(* IEC 61131-3 sources: trust-platform/crates/trust-runtime/tests/fixtures/control_pid/src, 10 files *)

(* ---- advanced_control_tests.st ---- *)
USING Control;

TEST_PROGRAM control_smith_predictor_models_delay_and_anchors_prediction_to_measurement
VAR
    Predictor : SmithPredictorFOPDT;
    Parameters : SmithPredictorParameters;
    State : SmithPredictorInitialState;
    Input : SmithPredictorInput;
    Output : SmithPredictorOutput;
    Accepted : BOOL;
END_VAR
Parameters.ProcessGain := LREAL#2.0;
Parameters.TimeConstant := LREAL#1.0;
Parameters.DeadTime := LREAL#1.0;
Parameters.OperatingOutput := LREAL#10.0;
Parameters.MaximumCorrection := LREAL#0.5;
Accepted := Predictor.Configure(Parameters := Parameters);
ASSERT_TRUE(Accepted);
State.ModelOutput := LREAL#10.0;
State.ProcessValue := LREAL#10.0;
Predictor.Initialize(State := State);
Input.ManipulatedValue := LREAL#1.0;
Input.ProcessValue := LREAL#10.0;
Input.CycleTime := LREAL#0.5;
Input.Enabled := TRUE;
Output := Predictor.Update(Input := Input);
ASSERT_TRUE(Output.Active);
ASSERT_TRUE(Output.HistoryComplete);
ASSERT_NEAR(EXPECTED := LREAL#10.8, ACTUAL := Output.DelayFreeModel, DELTA := LREAL#1.0e-12);
ASSERT_NEAR(EXPECTED := LREAL#10.0, ACTUAL := Output.DelayedModel, DELTA := LREAL#1.0e-12);
ASSERT_NEAR(EXPECTED := LREAL#10.8, ACTUAL := Output.PredictedProcessValue, DELTA := LREAL#1.0e-12);

Input.ProcessValue := LREAL#12.0;
Output := Predictor.Update(Input := Input);
ASSERT_NEAR(EXPECTED := LREAL#0.5, ACTUAL := Output.Correction, DELTA := LREAL#1.0e-12);
ASSERT_NEAR(EXPECTED := LREAL#11.78, ACTUAL := Output.PredictedProcessValue, DELTA := LREAL#1.0e-12);

Input.Enabled := FALSE;
Input.ProcessValue := LREAL#9.25;
Output := Predictor.Update(Input := Input);
ASSERT_FALSE(Output.Active);
ASSERT_NEAR(EXPECTED := LREAL#9.25, ACTUAL := Output.PredictedProcessValue, DELTA := LREAL#1.0e-12);

Parameters.TimeConstant := LREAL#0.0;
Accepted := Predictor.Configure(Parameters := Parameters);
ASSERT_FALSE(Accepted);
END_TEST_PROGRAM

TEST_PROGRAM control_pid_form_conversion_is_explicit_reversible_and_fail_closed
VAR
    Input : PIDFormParameters;
    Result : PIDFormConversionResult;
    Parallel : PIDFormParameters;
END_VAR

Input.Form := PIDParameterForm#Ideal;
Input.Proportional := LREAL#2.0;
Input.Integral := LREAL#10.0;
Input.Derivative := LREAL#0.5;
Result := ConvertPIDForm(Input := Input, Target := PIDParameterForm#Parallel);
ASSERT_TRUE(Result.Status = PIDFormConversionStatus#Valid);
ASSERT_NEAR(EXPECTED := LREAL#2.0, ACTUAL := Result.Parameters.Proportional, DELTA := LREAL#1.0e-12);
ASSERT_NEAR(EXPECTED := LREAL#0.2, ACTUAL := Result.Parameters.Integral, DELTA := LREAL#1.0e-12);
ASSERT_NEAR(EXPECTED := LREAL#1.0, ACTUAL := Result.Parameters.Derivative, DELTA := LREAL#1.0e-12);

Input.Form := PIDParameterForm#Series;
Result := ConvertPIDForm(Input := Input, Target := PIDParameterForm#Parallel);
ASSERT_TRUE(Result.Status = PIDFormConversionStatus#Valid);
ASSERT_NEAR(EXPECTED := LREAL#2.1, ACTUAL := Result.Parameters.Proportional, DELTA := LREAL#1.0e-12);
ASSERT_NEAR(EXPECTED := LREAL#0.2, ACTUAL := Result.Parameters.Integral, DELTA := LREAL#1.0e-12);
ASSERT_NEAR(EXPECTED := LREAL#1.0, ACTUAL := Result.Parameters.Derivative, DELTA := LREAL#1.0e-12);
Parallel := Result.Parameters;
Result := ConvertPIDForm(Input := Parallel, Target := PIDParameterForm#Series);
ASSERT_TRUE(Result.Status = PIDFormConversionStatus#Valid);
ASSERT_NEAR(EXPECTED := LREAL#2.0, ACTUAL := Result.Parameters.Proportional, DELTA := LREAL#1.0e-12);
ASSERT_NEAR(EXPECTED := LREAL#10.0, ACTUAL := Result.Parameters.Integral, DELTA := LREAL#1.0e-12);
ASSERT_NEAR(EXPECTED := LREAL#0.5, ACTUAL := Result.Parameters.Derivative, DELTA := LREAL#1.0e-12);

Parallel.Form := PIDParameterForm#Parallel;
Parallel.Proportional := LREAL#-2.0;
Parallel.Integral := LREAL#-0.2;
Parallel.Derivative := LREAL#-1.0;
Result := ConvertPIDForm(Input := Parallel, Target := PIDParameterForm#Ideal);
ASSERT_TRUE(Result.Status = PIDFormConversionStatus#Valid);
ASSERT_NEAR(EXPECTED := LREAL#-2.0, ACTUAL := Result.Parameters.Proportional, DELTA := LREAL#1.0e-12);
ASSERT_NEAR(EXPECTED := LREAL#10.0, ACTUAL := Result.Parameters.Integral, DELTA := LREAL#1.0e-12);
ASSERT_NEAR(EXPECTED := LREAL#0.5, ACTUAL := Result.Parameters.Derivative, DELTA := LREAL#1.0e-12);

Result := ConvertPIDForm(Input := Parallel, Target := PIDParameterForm#Parallel);
ASSERT_TRUE(Result.Status = PIDFormConversionStatus#Valid);
ASSERT_NEAR(EXPECTED := Parallel.Proportional, ACTUAL := Result.Parameters.Proportional, DELTA := LREAL#1.0e-12);

Input.Form := PIDParameterForm#Ideal;
Input.Proportional := LREAL#2.0;
Input.Integral := LREAL#0.0;
Input.Derivative := LREAL#0.5;
Result := ConvertPIDForm(Input := Input, Target := PIDParameterForm#Parallel);
ASSERT_TRUE(Result.Status = PIDFormConversionStatus#InvalidDomain);

Parallel.Form := PIDParameterForm#Parallel;
Parallel.Proportional := LREAL#1.0;
Parallel.Integral := LREAL#1.0;
Parallel.Derivative := LREAL#1.0;
Result := ConvertPIDForm(Input := Parallel, Target := PIDParameterForm#Series);
ASSERT_TRUE(Result.Status = PIDFormConversionStatus#NonRepresentable);
END_TEST_PROGRAM

TEST_PROGRAM control_smith_predictor_initialization_sets_the_correction_from_the_measurement
VAR
    Predictor : SmithPredictorFOPDT;
    State : SmithPredictorInitialState;
    Input : SmithPredictorInput;
    Output : SmithPredictorOutput;
END_VAR
(* Spec 37 §2.3: Initialize sets the initial correction from ProcessValue - ModelOutput. Before
   configuration no model interval runs, so the update reports that correction while it returns
   the measurement. *)
State.ModelOutput := LREAL#10.0;
State.ProcessValue := LREAL#12.0;
Predictor.Initialize(State := State);
Input.ProcessValue := LREAL#12.0;
Input.CycleTime := LREAL#0.5;
Input.Enabled := TRUE;
Output := Predictor.Update(Input := Input);
ASSERT_FALSE(Output.Active);
ASSERT_NEAR(EXPECTED := LREAL#12.0, ACTUAL := Output.PredictedProcessValue, DELTA := LREAL#1.0e-12);
ASSERT_NEAR(EXPECTED := LREAL#2.0, ACTUAL := Output.Correction, DELTA := LREAL#1.0e-12);
END_TEST_PROGRAM

TEST_PROGRAM control_smith_predictor_zero_delay_reduces_to_measurement
VAR
    Predictor : SmithPredictorFOPDT;
    Parameters : SmithPredictorParameters;
    State : SmithPredictorInitialState;
    Input : SmithPredictorInput;
    Output : SmithPredictorOutput;
END_VAR
Parameters.ProcessGain := LREAL#1.0;
Parameters.TimeConstant := LREAL#2.0;
Parameters.DeadTime := LREAL#0.0;
ASSERT_TRUE(Predictor.Configure(Parameters := Parameters));
Predictor.Initialize(State := State);
Input.ManipulatedValue := LREAL#4.0;
Input.ProcessValue := LREAL#7.25;
Input.CycleTime := LREAL#0.1;
Input.Enabled := TRUE;
Output := Predictor.Update(Input := Input);
ASSERT_NEAR(EXPECTED := LREAL#7.25, ACTUAL := Output.PredictedProcessValue, DELTA := LREAL#1.0e-12);
END_TEST_PROGRAM

TEST_PROGRAM control_pid_gain_scheduler_interpolates_tuning_and_preserves_common_policy
VAR
    Scheduler : PIDGainScheduler;
    Parameters : PIDGainScheduleParameters;
    Output : PIDGainScheduleOutput;
    Accepted : BOOL;
END_VAR
Parameters.PointCount := DINT#3;
Parameters.Points[0].OperatingPoint := LREAL#0.0;
Parameters.Points[0].Tuning.ProportionalGain := LREAL#1.0;
Parameters.Points[0].Tuning.IntegralGain := LREAL#0.1;
Parameters.Points[0].Tuning.DerivativeGain := LREAL#0.2;
Parameters.Points[0].Tuning.ProportionalSetpointWeight := LREAL#0.3;
Parameters.Points[0].Tuning.DerivativeSetpointWeight := LREAL#0.4;
Parameters.Points[0].Tuning.TrackingTime := LREAL#1.0;
Parameters.Points[1].OperatingPoint := LREAL#10.0;
Parameters.Points[1].Tuning.ProportionalGain := LREAL#2.0;
Parameters.Points[1].Tuning.IntegralGain := LREAL#0.2;
Parameters.Points[1].Tuning.DerivativeGain := LREAL#0.4;
Parameters.Points[1].Tuning.ProportionalSetpointWeight := LREAL#0.5;
Parameters.Points[1].Tuning.DerivativeSetpointWeight := LREAL#0.6;
Parameters.Points[1].Tuning.TrackingTime := LREAL#2.0;
Parameters.Points[2].OperatingPoint := LREAL#20.0;
Parameters.Points[2].Tuning.ProportionalGain := LREAL#4.0;
Parameters.Points[2].Tuning.IntegralGain := LREAL#0.4;
Parameters.Points[2].Tuning.DerivativeGain := LREAL#0.8;
Parameters.Points[2].Tuning.ProportionalSetpointWeight := LREAL#0.7;
Parameters.Points[2].Tuning.DerivativeSetpointWeight := LREAL#0.8;
Parameters.Points[2].Tuning.TrackingTime := LREAL#4.0;
Parameters.CommonParameters.Bias := LREAL#12.0;
Parameters.CommonParameters.OutputMinimum := LREAL#0.0;
Parameters.CommonParameters.OutputMaximum := LREAL#100.0;
Parameters.CommonParameters.RateMinimum := LREAL#-5.0;
Parameters.CommonParameters.RateMaximum := LREAL#7.0;
Parameters.CommonParameters.AntiWindup := PIDAntiWindup#Combined;
Accepted := Scheduler.Configure(Parameters := Parameters);
ASSERT_TRUE(Accepted);
Scheduler.Initialize(OperatingPoint := LREAL#5.0);
Output := Scheduler.Update(OperatingPoint := LREAL#5.0, CycleTime := LREAL#0.1);
ASSERT_TRUE(Output.Valid);
ASSERT_FALSE(Output.Clamped);
ASSERT_TRUE(Output.LowerIndex = DINT#0);
ASSERT_TRUE(Output.UpperIndex = DINT#1);
ASSERT_NEAR(EXPECTED := LREAL#0.5, ACTUAL := Output.Fraction, DELTA := LREAL#1.0e-12);
ASSERT_NEAR(EXPECTED := LREAL#1.5, ACTUAL := Output.Parameters.ProportionalGain, DELTA := LREAL#1.0e-12);
ASSERT_NEAR(EXPECTED := LREAL#0.15, ACTUAL := Output.Parameters.IntegralGain, DELTA := LREAL#1.0e-12);
ASSERT_NEAR(EXPECTED := LREAL#0.3, ACTUAL := Output.Parameters.DerivativeGain, DELTA := LREAL#1.0e-12);
ASSERT_NEAR(EXPECTED := LREAL#0.4, ACTUAL := Output.Parameters.ProportionalSetpointWeight, DELTA := LREAL#1.0e-12);
ASSERT_NEAR(EXPECTED := LREAL#0.5, ACTUAL := Output.Parameters.DerivativeSetpointWeight, DELTA := LREAL#1.0e-12);
ASSERT_NEAR(EXPECTED := LREAL#1.5, ACTUAL := Output.Parameters.TrackingTime, DELTA := LREAL#1.0e-12);
ASSERT_NEAR(EXPECTED := LREAL#12.0, ACTUAL := Output.Parameters.Bias, DELTA := LREAL#1.0e-12);
ASSERT_NEAR(EXPECTED := LREAL#100.0, ACTUAL := Output.Parameters.OutputMaximum, DELTA := LREAL#1.0e-12);
ASSERT_TRUE(Output.Parameters.AntiWindup = PIDAntiWindup#Combined);

Output := Scheduler.Update(OperatingPoint := LREAL#-5.0, CycleTime := LREAL#0.1);
ASSERT_TRUE(Output.Clamped);
ASSERT_NEAR(EXPECTED := LREAL#1.0, ACTUAL := Output.Parameters.ProportionalGain, DELTA := LREAL#1.0e-12);

Parameters.Points[1].OperatingPoint := LREAL#0.0;
Accepted := Scheduler.Configure(Parameters := Parameters);
ASSERT_FALSE(Accepted);
Output := Scheduler.Update(OperatingPoint := LREAL#15.0, CycleTime := LREAL#0.1);
ASSERT_NEAR(EXPECTED := LREAL#3.0, ACTUAL := Output.Parameters.ProportionalGain, DELTA := LREAL#1.0e-12);
END_TEST_PROGRAM

TEST_PROGRAM control_pid_gain_scheduler_filters_the_operating_point
VAR
    Scheduler : PIDGainScheduler;
    Parameters : PIDGainScheduleParameters;
    Output : PIDGainScheduleOutput;
END_VAR
Parameters.PointCount := DINT#2;
Parameters.Points[0].OperatingPoint := LREAL#0.0;
Parameters.Points[0].Tuning.ProportionalGain := LREAL#1.0;
Parameters.Points[0].Tuning.TrackingTime := LREAL#1.0;
Parameters.Points[1].OperatingPoint := LREAL#10.0;
Parameters.Points[1].Tuning.ProportionalGain := LREAL#3.0;
Parameters.Points[1].Tuning.TrackingTime := LREAL#1.0;
Parameters.CommonParameters.OutputMinimum := LREAL#-100.0;
Parameters.CommonParameters.OutputMaximum := LREAL#100.0;
Parameters.CommonParameters.RateMinimum := LREAL#-100.0;
Parameters.CommonParameters.RateMaximum := LREAL#100.0;
Parameters.FilterTimeConstant := LREAL#1.0;
ASSERT_TRUE(Scheduler.Configure(Parameters := Parameters));
Scheduler.Initialize(OperatingPoint := LREAL#0.0);
Output := Scheduler.Update(OperatingPoint := LREAL#10.0, CycleTime := LREAL#1.0);
ASSERT_NEAR(EXPECTED := LREAL#5.0, ACTUAL := Output.FilteredOperatingPoint, DELTA := LREAL#1.0e-12);
ASSERT_NEAR(EXPECTED := LREAL#2.0, ACTUAL := Output.Parameters.ProportionalGain, DELTA := LREAL#1.0e-12);
END_TEST_PROGRAM

TEST_PROGRAM control_static_decoupler_maps_and_recovers_two_channel_commands
VAR
    Decoupler : StaticDecoupler2x2;
    Parameters : StaticDecoupler2x2Parameters;
    VirtualCommand : ControlVector2;
    ActuatorCommand : ControlVector2;
    Recovered : ControlVector2;
    Status : StaticDecoupler2x2Status;
    Accepted : BOOL;
END_VAR
VirtualCommand.First := LREAL#3.0;
ActuatorCommand := Decoupler.ToActuators(VirtualCommand := VirtualCommand);
ASSERT_NEAR(EXPECTED := LREAL#0.0, ACTUAL := ActuatorCommand.First, DELTA := LREAL#1.0e-12);
ASSERT_NEAR(EXPECTED := LREAL#0.0, ACTUAL := ActuatorCommand.Second, DELTA := LREAL#1.0e-12);

Parameters.GainMatrix.G11 := LREAL#2.0;
Parameters.GainMatrix.G12 := LREAL#1.0;
Parameters.GainMatrix.G21 := LREAL#1.0;
Parameters.GainMatrix.G22 := LREAL#2.0;
Parameters.ActuatorBias.First := LREAL#10.0;
Parameters.ActuatorBias.Second := LREAL#20.0;
Parameters.SingularityTolerance := LREAL#1.0e-9;
Accepted := Decoupler.Configure(Parameters := Parameters);
ASSERT_TRUE(Accepted);
Status := Decoupler.Snapshot();
ASSERT_TRUE(Status.Configured);
ASSERT_NEAR(EXPECTED := LREAL#3.0, ACTUAL := Status.Determinant, DELTA := LREAL#1.0e-12);
ActuatorCommand := Decoupler.ToActuators(VirtualCommand := VirtualCommand);
ASSERT_NEAR(EXPECTED := LREAL#12.0, ACTUAL := ActuatorCommand.First, DELTA := LREAL#1.0e-12);
ASSERT_NEAR(EXPECTED := LREAL#19.0, ACTUAL := ActuatorCommand.Second, DELTA := LREAL#1.0e-12);
Recovered := Decoupler.ToVirtual(ActuatorCommand := ActuatorCommand);
ASSERT_NEAR(EXPECTED := LREAL#3.0, ACTUAL := Recovered.First, DELTA := LREAL#1.0e-12);
ASSERT_NEAR(EXPECTED := LREAL#0.0, ACTUAL := Recovered.Second, DELTA := LREAL#1.0e-12);

Parameters.GainMatrix.G11 := LREAL#1000000.0;
Parameters.GainMatrix.G12 := LREAL#1000000.0;
Parameters.GainMatrix.G21 := LREAL#1000000.0;
Parameters.GainMatrix.G22 := LREAL#1000000.01;
Parameters.SingularityTolerance := LREAL#1.0e-6;
Accepted := Decoupler.Configure(Parameters := Parameters);
ASSERT_FALSE(Accepted);
ActuatorCommand := Decoupler.ToActuators(VirtualCommand := VirtualCommand);
ASSERT_NEAR(EXPECTED := LREAL#12.0, ACTUAL := ActuatorCommand.First, DELTA := LREAL#1.0e-12);
ASSERT_NEAR(EXPECTED := LREAL#19.0, ACTUAL := ActuatorCommand.Second, DELTA := LREAL#1.0e-12);

Parameters.GainMatrix.G11 := LREAL#1.0;
Parameters.GainMatrix.G12 := LREAL#2.0;
Parameters.GainMatrix.G21 := LREAL#2.0;
Parameters.GainMatrix.G22 := LREAL#4.0;
Accepted := Decoupler.Configure(Parameters := Parameters);
ASSERT_FALSE(Accepted);
ActuatorCommand := Decoupler.ToActuators(VirtualCommand := VirtualCommand);
ASSERT_NEAR(EXPECTED := LREAL#12.0, ACTUAL := ActuatorCommand.First, DELTA := LREAL#1.0e-12);
ASSERT_NEAR(EXPECTED := LREAL#19.0, ACTUAL := ActuatorCommand.Second, DELTA := LREAL#1.0e-12);
END_TEST_PROGRAM

(* ---- antiwindup_tests.st ---- *)
USING Control;

TEST_PROGRAM control_pid_back_calculation_and_clamping_retain_distinct_nominal_states
VAR
    BackCalculationController : PID;
    ClampingController : PID;
    Parameters : PIDParameters;
    InitialState : PIDInitialState;
    Input : PIDInput;
    Output : LREAL;
END_VAR

Parameters.IntegralGain := LREAL#4.0;
Parameters.OutputMinimum := LREAL#0.0;
Parameters.OutputMaximum := LREAL#3.0;
Parameters.RateMinimum := LREAL#-1000.0;
Parameters.RateMaximum := LREAL#1000.0;
Parameters.TrackingTime := LREAL#2.0;
BackCalculationController.Configure(Parameters := Parameters);
BackCalculationController.Initialize(State := InitialState);

Input.Setpoint := LREAL#1.0;
Input.CycleTime := LREAL#1.0;
Output := BackCalculationController.Update(Input := Input);
ASSERT_NEAR(EXPECTED := LREAL#3.0, ACTUAL := Output, DELTA := LREAL#3.0e-12);
Input.Setpoint := LREAL#-0.125;
Output := BackCalculationController.Update(Input := Input);
ASSERT_NEAR(EXPECTED := LREAL#3.0, ACTUAL := Output, DELTA := LREAL#3.0e-12);

Parameters.TrackingTime := LREAL#1.0;
ClampingController.Configure(Parameters := Parameters);
ClampingController.Initialize(State := InitialState);
Input.Setpoint := LREAL#1.0;
Output := ClampingController.Update(Input := Input);
ASSERT_NEAR(EXPECTED := LREAL#3.0, ACTUAL := Output, DELTA := LREAL#3.0e-12);
Input.Setpoint := LREAL#-0.125;
Output := ClampingController.Update(Input := Input);
ASSERT_NEAR(EXPECTED := LREAL#2.5, ACTUAL := Output, DELTA := LREAL#2.5e-12);
END_TEST_PROGRAM

TEST_PROGRAM control_pid_combined_anti_windup_allows_integration_away_from_saturation
VAR
    Controller : PID;
    Parameters : PIDParameters;
    InitialState : PIDInitialState;
    Input : PIDInput;
    Output : LREAL;
END_VAR

Parameters.IntegralGain := LREAL#1.0;
Parameters.OutputMinimum := LREAL#0.0;
Parameters.OutputMaximum := LREAL#3.0;
Parameters.RateMinimum := LREAL#-1000.0;
Parameters.RateMaximum := LREAL#1000.0;
Parameters.TrackingTime := LREAL#2.0;
Parameters.AntiWindup := PIDAntiWindup#Combined;
InitialState.NominalOutput := LREAL#4.0;
InitialState.SaturatedOutput := LREAL#3.0;
Controller.Configure(Parameters := Parameters);
Controller.Initialize(State := InitialState);

Input.Setpoint := LREAL#1.0;
Input.CycleTime := LREAL#1.0;
Output := Controller.Update(Input := Input);
ASSERT_NEAR(EXPECTED := LREAL#3.0, ACTUAL := Output, DELTA := LREAL#3.0e-12);

Input.Setpoint := LREAL#-0.75;
Output := Controller.Update(Input := Input);
ASSERT_NEAR(EXPECTED := LREAL#2.75, ACTUAL := Output, DELTA := LREAL#2.75e-12);
END_TEST_PROGRAM

(* ---- configuration_tests.st ---- *)
(* Specification 45 sections 2.4/2.5 and 3.2/3.3: complete value-copy configuration,
   retained histories, and initialization without an update. *)
USING Control;

TEST_PROGRAM control_pid_configuration_copies_parameters_and_preserves_every_history
VAR
    Controller : PID;
    Parameters : PIDParameters;
    AcceptedParameters : PIDParameters;
    InitialState : PIDInitialState;
    ZeroState : PIDInitialState;
    Observed : PIDInitialState;
    Input : PIDInput;
    Output : LREAL;
END_VAR

InitialState.Setpoint := LREAL#10.0;
InitialState.SetpointRate := LREAL#2.0;
InitialState.ProcessValue := LREAL#8.0;
InitialState.ProcessValueRate := LREAL#-1.0;
InitialState.FeedForward := LREAL#3.0;
InitialState.NominalOutput := LREAL#20.0;
InitialState.SaturatedOutput := LREAL#19.0;
Parameters.OutputMinimum := LREAL#-100.0;
Parameters.OutputMaximum := LREAL#100.0;
Parameters.RateMinimum := LREAL#-1000.0;
Parameters.RateMaximum := LREAL#1000.0;
Parameters.TrackingTime := LREAL#1.0;
Controller.Configure(Parameters := Parameters);
Controller.Initialize(State := InitialState);
Observed := Controller.GetState();
ASSERT_NEAR(EXPECTED := LREAL#10.0, ACTUAL := Observed.Setpoint, DELTA := LREAL#1.0e-12);
ASSERT_NEAR(EXPECTED := LREAL#2.0, ACTUAL := Observed.SetpointRate, DELTA := LREAL#1.0e-12);
ASSERT_NEAR(EXPECTED := LREAL#8.0, ACTUAL := Observed.ProcessValue, DELTA := LREAL#1.0e-12);
ASSERT_NEAR(EXPECTED := LREAL#-1.0, ACTUAL := Observed.ProcessValueRate, DELTA := LREAL#1.0e-12);
ASSERT_NEAR(EXPECTED := LREAL#3.0, ACTUAL := Observed.FeedForward, DELTA := LREAL#1.0e-12);
ASSERT_NEAR(EXPECTED := LREAL#20.0, ACTUAL := Observed.NominalOutput, DELTA := LREAL#1.0e-12);
ASSERT_NEAR(EXPECTED := LREAL#19.0, ACTUAL := Observed.SaturatedOutput, DELTA := LREAL#1.0e-12);

Parameters.ProportionalGain := LREAL#2.0;
Parameters.IntegralGain := LREAL#0.5;
Parameters.DerivativeGain := LREAL#0.25;
Parameters.ProportionalSetpointWeight := LREAL#0.4;
Parameters.DerivativeSetpointWeight := LREAL#0.3;
Parameters.Bias := LREAL#7.0;
Parameters.OutputMinimum := LREAL#-30.0;
Parameters.OutputMaximum := LREAL#40.0;
Parameters.RateMinimum := LREAL#-4.0;
Parameters.RateMaximum := LREAL#6.0;
Parameters.TrackingTime := LREAL#2.0;
Parameters.AntiWindup := PIDAntiWindup#Combined;
Controller.Configure(Parameters := Parameters);
Observed := Controller.GetState();
ASSERT_NEAR(EXPECTED := LREAL#10.0, ACTUAL := Observed.Setpoint, DELTA := LREAL#1.0e-12);
ASSERT_NEAR(EXPECTED := LREAL#2.0, ACTUAL := Observed.SetpointRate, DELTA := LREAL#1.0e-12);
ASSERT_NEAR(EXPECTED := LREAL#8.0, ACTUAL := Observed.ProcessValue, DELTA := LREAL#1.0e-12);
ASSERT_NEAR(EXPECTED := LREAL#-1.0, ACTUAL := Observed.ProcessValueRate, DELTA := LREAL#1.0e-12);
ASSERT_NEAR(EXPECTED := LREAL#3.0, ACTUAL := Observed.FeedForward, DELTA := LREAL#1.0e-12);
ASSERT_NEAR(EXPECTED := LREAL#20.0, ACTUAL := Observed.NominalOutput, DELTA := LREAL#1.0e-12);
ASSERT_NEAR(EXPECTED := LREAL#19.0, ACTUAL := Observed.SaturatedOutput, DELTA := LREAL#1.0e-12);

(* Mutating the caller's record after Configure cannot alter the accepted copy. *)
AcceptedParameters := Parameters;
Parameters.ProportionalGain := LREAL#100.0;
Parameters.IntegralGain := LREAL#0.0;
Parameters.DerivativeGain := LREAL#0.0;
Parameters.ProportionalSetpointWeight := LREAL#1.0;
Parameters.DerivativeSetpointWeight := LREAL#1.0;
Parameters.Bias := LREAL#-10.0;
Parameters.OutputMinimum := LREAL#-100.0;
Parameters.OutputMaximum := LREAL#100.0;
Parameters.RateMinimum := LREAL#-1000.0;
Parameters.RateMaximum := LREAL#1000.0;
Parameters.TrackingTime := LREAL#10.0;
Parameters.AntiWindup := PIDAntiWindup#BackCalculation;

Input.Setpoint := LREAL#12.0;
Input.ProcessValue := LREAL#9.0;
Input.FeedForward := LREAL#5.0;
Input.CycleTime := LREAL#0.5;
Output := Controller.Update(Input := Input);
(* 20 - 0.4 + 0.75 - 0.6 + 2 = 21.75; rate interval is [17,22]. *)
ASSERT_NEAR(EXPECTED := LREAL#21.75, ACTUAL := Output, DELTA := LREAL#1.0e-10);
Input.Setpoint := LREAL#13.0;
Input.ProcessValue := LREAL#11.0;
Input.FeedForward := LREAL#6.0;
Input.CycleTime := LREAL#0.25;
Output := Controller.Update(Input := Input);
Observed := Controller.GetState();
ASSERT_NEAR(EXPECTED := LREAL#20.75, ACTUAL := Output, DELTA := LREAL#1.0e-10);
ASSERT_NEAR(EXPECTED := LREAL#18.60625, ACTUAL := Observed.NominalOutput, DELTA := LREAL#1.0e-10);
ASSERT_NEAR(EXPECTED := LREAL#4.0, ACTUAL := Observed.SetpointRate, DELTA := LREAL#1.0e-12);
ASSERT_NEAR(EXPECTED := LREAL#8.0, ACTUAL := Observed.ProcessValueRate, DELTA := LREAL#1.0e-12);

Input.Mode := PIDMode#Manual;
Input.ManualOutput := LREAL#100.0;
Input.CycleTime := LREAL#10.0;
ASSERT_NEAR(EXPECTED := LREAL#40.0, ACTUAL := Controller.Update(Input := Input), DELTA := LREAL#1.0e-12);
Input.ManualOutput := LREAL#-100.0;
Input.CycleTime := LREAL#20.0;
ASSERT_NEAR(EXPECTED := LREAL#-30.0, ACTUAL := Controller.Update(Input := Input), DELTA := LREAL#1.0e-12);
Input.ManualOutput := LREAL#100.0;
Input.CycleTime := LREAL#0.5;
ASSERT_NEAR(EXPECTED := LREAL#-27.0, ACTUAL := Controller.Update(Input := Input), DELTA := LREAL#1.0e-12);

Controller.Initialize(State := ZeroState);
Input.Mode := PIDMode#Auto;
Input.Setpoint := LREAL#100.0;
Input.ProcessValue := LREAL#0.0;
Input.FeedForward := LREAL#0.0;
Input.CycleTime := LREAL#1.0;
Output := Controller.Update(Input := Input);
Observed := Controller.GetState();
(* Combined removes 50 of the 131.5 saturation error, then back-calculates
   with coefficient 1/2: 137.5 - 50 - (87.5 - 6)/2 = 46.75. *)
ASSERT_NEAR(EXPECTED := LREAL#6.0, ACTUAL := Output, DELTA := LREAL#1.0e-12);
ASSERT_NEAR(EXPECTED := LREAL#46.75, ACTUAL := Observed.NominalOutput, DELTA := LREAL#1.0e-10);

(* The same complete record's Bias takes effect when integral action is zero. *)
Parameters := AcceptedParameters;
Parameters.IntegralGain := LREAL#0.0;
Controller.Configure(Parameters := Parameters);
Parameters.Bias := LREAL#700.0;
Controller.Initialize(State := ZeroState);
Input.Setpoint := LREAL#0.0;
Input.CycleTime := LREAL#2.0;
ASSERT_NEAR(EXPECTED := LREAL#7.0, ACTUAL := Controller.Update(Input := Input), DELTA := LREAL#1.0e-12);
END_TEST_PROGRAM

(* Specification 45 sections 4.2/4.3 and 6: separate filter histories continue
   across reconfiguration, using each call's own elapsed interval. *)
TEST_PROGRAM control_low_pass_reconfiguration_preserves_both_stages_and_actual_intervals
VAR
    Filter : LowPass;
    Parameters : LowPassParameters;
END_VAR
Parameters.TimeConstant := LREAL#1.5;
Parameters.Order := FilterOrder#SecondOrder;
Filter.Configure(Parameters := Parameters);
Filter.Initialize(Input := LREAL#2.0);
ASSERT_NEAR(EXPECTED := LREAL#2.5, ACTUAL := Filter.Update(Input := LREAL#4.0, CycleTime := LREAL#1.0), DELTA := LREAL#1.0e-12);

Parameters.TimeConstant := LREAL#0.75;
Filter.Configure(Parameters := Parameters);
Parameters.TimeConstant := LREAL#100.0;
Parameters.Order := FilterOrder#FirstOrder;
ASSERT_NEAR(EXPECTED := LREAL#3.0, ACTUAL := Filter.Update(Input := LREAL#4.0, CycleTime := LREAL#0.5), DELTA := LREAL#1.0e-12);

Parameters.TimeConstant := LREAL#0.75;
Filter.Configure(Parameters := Parameters);
ASSERT_NEAR(EXPECTED := LREAL#4.25, ACTUAL := Filter.Update(Input := LREAL#5.0, CycleTime := LREAL#0.5), DELTA := LREAL#1.0e-12);
Parameters.Order := FilterOrder#SecondOrder;
Filter.Configure(Parameters := Parameters);
ASSERT_NEAR(EXPECTED := LREAL#3.8125, ACTUAL := Filter.Update(Input := LREAL#5.0, CycleTime := LREAL#0.5), DELTA := LREAL#1.0e-12);
END_TEST_PROGRAM

(* ---- filter_tests.st ---- *)
USING Control;

TEST_PROGRAM control_low_pass_matches_listing_four_for_both_orders
VAR
    FirstOrderFilter : LowPass;
    SecondOrderFilter : LowPass;
    Parameters : LowPassParameters;
    Output : LREAL;
END_VAR

Parameters.TimeConstant := LREAL#1.5;
FirstOrderFilter.Configure(Parameters := Parameters);
FirstOrderFilter.Initialize(Input := LREAL#2.0);
Output := FirstOrderFilter.Update(Input := LREAL#4.0, CycleTime := LREAL#1.0);
ASSERT_NEAR(EXPECTED := LREAL#3.0, ACTUAL := Output, DELTA := LREAL#3.0e-12);

Parameters.Order := FilterOrder#SecondOrder;
SecondOrderFilter.Configure(Parameters := Parameters);
SecondOrderFilter.Initialize(Input := LREAL#2.0);
Output := SecondOrderFilter.Update(Input := LREAL#4.0, CycleTime := LREAL#1.0);
ASSERT_NEAR(EXPECTED := LREAL#2.5, ACTUAL := Output, DELTA := LREAL#2.5e-12);
Output := SecondOrderFilter.Update(Input := LREAL#4.0, CycleTime := LREAL#1.0);
ASSERT_NEAR(EXPECTED := LREAL#3.0, ACTUAL := Output, DELTA := LREAL#3.0e-12);

Parameters.TimeConstant := LREAL#0.5;
Parameters.Order := FilterOrder#FirstOrder;
FirstOrderFilter.Configure(Parameters := Parameters);
FirstOrderFilter.Initialize(Input := LREAL#2.0);
Output := FirstOrderFilter.Update(Input := LREAL#4.0, CycleTime := LREAL#1.0);
ASSERT_NEAR(EXPECTED := LREAL#4.0, ACTUAL := Output, DELTA := LREAL#4.0e-12);

Parameters.Order := FilterOrder#SecondOrder;
SecondOrderFilter.Configure(Parameters := Parameters);
SecondOrderFilter.Initialize(Input := LREAL#2.0);
Output := SecondOrderFilter.Update(Input := LREAL#4.0, CycleTime := LREAL#1.0);
ASSERT_NEAR(EXPECTED := LREAL#4.0, ACTUAL := Output, DELTA := LREAL#4.0e-12);
END_TEST_PROGRAM

(* ---- instance_tests.st ---- *)
USING Control;

TEST_PROGRAM control_pid_and_filter_histories_are_instance_local
VAR
    PidA : PID;
    PidB : PID;
    PidAAlone : PID;
    PidBAlone : PID;
    PidParametersA : PIDParameters;
    PidParametersB : PIDParameters;
    PidStateA : PIDInitialState;
    PidStateB : PIDInitialState;
    PidInputA : PIDInput;
    PidInputB : PIDInput;
    A1 : LREAL;
    A2 : LREAL;
    B1 : LREAL;
    B2 : LREAL;
    FilterA : LowPass;
    FilterB : LowPass;
    FilterAAlone : LowPass;
    FilterBAlone : LowPass;
    FilterParametersA : LowPassParameters;
    FilterParametersB : LowPassParameters;
    FA1 : LREAL;
    FA2 : LREAL;
    FB1 : LREAL;
    FB2 : LREAL;
END_VAR

PidParametersA.ProportionalGain := LREAL#1.0;
PidParametersA.IntegralGain := LREAL#1.0;
PidParametersA.ProportionalSetpointWeight := LREAL#0.5;
PidParametersA.OutputMinimum := LREAL#-100.0;
PidParametersA.OutputMaximum := LREAL#100.0;
PidParametersA.RateMinimum := LREAL#-1000.0;
PidParametersA.RateMaximum := LREAL#1000.0;
PidParametersA.TrackingTime := LREAL#1.0;
PidParametersB := PidParametersA;
PidParametersB.ProportionalGain := LREAL#2.0;
PidParametersB.IntegralGain := LREAL#0.5;
PidStateB.NominalOutput := LREAL#5.0;
PidStateB.SaturatedOutput := LREAL#5.0;

PidA.Configure(Parameters := PidParametersA);
PidA.Initialize(State := PidStateA);
PidAAlone.Configure(Parameters := PidParametersA);
PidAAlone.Initialize(State := PidStateA);
PidB.Configure(Parameters := PidParametersB);
PidB.Initialize(State := PidStateB);
PidBAlone.Configure(Parameters := PidParametersB);
PidBAlone.Initialize(State := PidStateB);

PidInputA.Setpoint := LREAL#1.0;
PidInputA.CycleTime := LREAL#0.1;
PidInputB.Setpoint := LREAL#-2.0;
PidInputB.ProcessValue := LREAL#0.5;
PidInputB.CycleTime := LREAL#0.2;
A1 := PidA.Update(Input := PidInputA);
B1 := PidB.Update(Input := PidInputB);
PidInputA.ProcessValue := LREAL#0.2;
A2 := PidA.Update(Input := PidInputA);
PidInputB.ProcessValue := LREAL#0.0;
B2 := PidB.Update(Input := PidInputB);

PidInputA.ProcessValue := LREAL#0.0;
ASSERT_NEAR(EXPECTED := A1, ACTUAL := PidAAlone.Update(Input := PidInputA), DELTA := LREAL#1.0e-12);
PidInputA.ProcessValue := LREAL#0.2;
ASSERT_NEAR(EXPECTED := A2, ACTUAL := PidAAlone.Update(Input := PidInputA), DELTA := LREAL#1.0e-12);

PidInputB.ProcessValue := LREAL#0.5;
ASSERT_NEAR(EXPECTED := B1, ACTUAL := PidBAlone.Update(Input := PidInputB), DELTA := LREAL#1.0e-12);
PidInputB.ProcessValue := LREAL#0.0;
ASSERT_NEAR(EXPECTED := B2, ACTUAL := PidBAlone.Update(Input := PidInputB), DELTA := LREAL#1.0e-12);

FilterParametersA.TimeConstant := LREAL#1.5;
FilterParametersB.TimeConstant := LREAL#2.5;
FilterParametersB.Order := FilterOrder#SecondOrder;
FilterA.Configure(Parameters := FilterParametersA);
FilterA.Initialize(Input := LREAL#0.0);
FilterAAlone.Configure(Parameters := FilterParametersA);
FilterAAlone.Initialize(Input := LREAL#0.0);
FilterB.Configure(Parameters := FilterParametersB);
FilterB.Initialize(Input := LREAL#10.0);
FilterBAlone.Configure(Parameters := FilterParametersB);
FilterBAlone.Initialize(Input := LREAL#10.0);

FA1 := FilterA.Update(Input := LREAL#4.0, CycleTime := LREAL#1.0);
FB1 := FilterB.Update(Input := LREAL#2.0, CycleTime := LREAL#0.5);
FA2 := FilterA.Update(Input := LREAL#6.0, CycleTime := LREAL#1.0);
FB2 := FilterB.Update(Input := LREAL#4.0, CycleTime := LREAL#0.5);

ASSERT_NEAR(EXPECTED := FA1, ACTUAL := FilterAAlone.Update(Input := LREAL#4.0, CycleTime := LREAL#1.0), DELTA := LREAL#1.0e-12);
ASSERT_NEAR(EXPECTED := FA2, ACTUAL := FilterAAlone.Update(Input := LREAL#6.0, CycleTime := LREAL#1.0), DELTA := LREAL#1.0e-12);
ASSERT_NEAR(EXPECTED := FB1, ACTUAL := FilterBAlone.Update(Input := LREAL#2.0, CycleTime := LREAL#0.5), DELTA := LREAL#1.0e-12);
ASSERT_NEAR(EXPECTED := FB2, ACTUAL := FilterBAlone.Update(Input := LREAL#4.0, CycleTime := LREAL#0.5), DELTA := LREAL#1.0e-12);
END_TEST_PROGRAM

(* ---- main.st ---- *)
PROGRAM Main
END_PROGRAM

(* ---- modes_tests.st ---- *)
USING Control;

TEST_PROGRAM control_pid_manual_limits_output_but_retains_nominal_history
VAR
    Controller : PID;
    Parameters : PIDParameters;
    InitialState : PIDInitialState;
    Input : PIDInput;
    Output : LREAL;
END_VAR

Parameters.IntegralGain := LREAL#1.0;
Parameters.OutputMinimum := LREAL#0.0;
Parameters.OutputMaximum := LREAL#10.0;
Parameters.RateMinimum := LREAL#-2.0;
Parameters.RateMaximum := LREAL#3.0;
Parameters.TrackingTime := LREAL#0.5;
InitialState.NominalOutput := LREAL#5.0;
InitialState.SaturatedOutput := LREAL#5.0;
Controller.Configure(Parameters := Parameters);
Controller.Initialize(State := InitialState);

Input.ManualOutput := LREAL#9.0;
Input.Mode := PIDMode#Manual;
Input.CycleTime := LREAL#0.5;
Output := Controller.Update(Input := Input);
ASSERT_NEAR(EXPECTED := LREAL#6.5, ACTUAL := Output, DELTA := LREAL#6.5e-12);

Input.Mode := PIDMode#Auto;
Output := Controller.Update(Input := Input);
ASSERT_NEAR(EXPECTED := LREAL#8.0, ACTUAL := Output, DELTA := LREAL#8.0e-12);
END_TEST_PROGRAM

TEST_PROGRAM control_pid_track_preloads_only_the_incremental_form
VAR
    IntegralController : PID;
    PositionalController : PID;
    Parameters : PIDParameters;
    InitialState : PIDInitialState;
    Input : PIDInput;
    Output : LREAL;
END_VAR

Parameters.ProportionalGain := LREAL#2.0;
Parameters.IntegralGain := LREAL#1.0;
Parameters.ProportionalSetpointWeight := LREAL#0.5;
Parameters.OutputMinimum := LREAL#-100.0;
Parameters.OutputMaximum := LREAL#100.0;
Parameters.RateMinimum := LREAL#-1000.0;
Parameters.RateMaximum := LREAL#1000.0;
Parameters.TrackingTime := LREAL#1.0;
IntegralController.Configure(Parameters := Parameters);
IntegralController.Initialize(State := InitialState);

Input.Setpoint := LREAL#1.0;
Input.TrackingOutput := LREAL#7.0;
Input.Mode := PIDMode#Track;
Input.CycleTime := LREAL#0.1;
Output := IntegralController.Update(Input := Input);
ASSERT_NEAR(EXPECTED := LREAL#8.1, ACTUAL := Output, DELTA := LREAL#8.1e-12);

Parameters.IntegralGain := LREAL#0.0;
Parameters.Bias := LREAL#1.0;
PositionalController.Configure(Parameters := Parameters);
PositionalController.Initialize(State := InitialState);
Output := PositionalController.Update(Input := Input);
ASSERT_NEAR(EXPECTED := LREAL#3.0, ACTUAL := Output, DELTA := LREAL#3.0e-12);
END_TEST_PROGRAM

(* ---- scenario_tests.st ---- *)
USING Control;

TEST_PROGRAM control_pid_replays_paper_example_1_manual_to_auto
VAR
    Controller : PID;
    Parameters : PIDParameters;
    State : PIDInitialState;
    Input : PIDInput;
    Output : LREAL;
END_VAR

Parameters.ProportionalGain := LREAL#0.6666666666666667;
Parameters.IntegralGain := LREAL#0.6666666666666667;
Parameters.ProportionalSetpointWeight := LREAL#1.0;
Parameters.OutputMinimum := LREAL#-1.0e100;
Parameters.OutputMaximum := LREAL#1.0e100;
Parameters.RateMinimum := LREAL#-1.0e100;
Parameters.RateMaximum := LREAL#1.0e100;
Parameters.TrackingTime := LREAL#1.0;
Controller.Configure(Parameters := Parameters);
Controller.Initialize(State := State);

Input.Setpoint := LREAL#3.0;
Input.CycleTime := LREAL#0.01;
Input.Mode := PIDMode#Manual;
Output := Controller.Update(Input := Input);
ASSERT_NEAR(EXPECTED := LREAL#0.0, ACTUAL := Output, DELTA := LREAL#1.0e-12);

Input.ManualOutput := LREAL#1.0;
Output := Controller.Update(Input := Input);
ASSERT_NEAR(EXPECTED := LREAL#1.0, ACTUAL := Output, DELTA := LREAL#1.0e-12);

(* Auto resumes from the nominal manual command retained by Listing 3. *)
Input.ProcessValue := LREAL#1.0;
Input.Mode := PIDMode#Auto;
Output := Controller.Update(Input := Input);
ASSERT_NEAR(EXPECTED := LREAL#0.3466666666666667, ACTUAL := Output, DELTA := LREAL#1.0e-12);

State.Setpoint := LREAL#3.0;
State.ProcessValue := LREAL#3.0;
State.NominalOutput := LREAL#3.0;
State.SaturatedOutput := LREAL#3.0;
Controller.Initialize(State := State);
Input.ProcessValue := LREAL#3.0;
Output := Controller.Update(Input := Input);
ASSERT_NEAR(EXPECTED := LREAL#3.0, ACTUAL := Output, DELTA := LREAL#1.0e-12);
END_TEST_PROGRAM

TEST_PROGRAM control_pid_replays_paper_example_2_form_switch_and_rate_limit
VAR
    Controller : PID;
    LimitedController : PID;
    Parameters : PIDParameters;
    State : PIDInitialState;
    Input : PIDInput;
    Output : LREAL;
END_VAR

Parameters.ProportionalGain := LREAL#0.6666666666666667;
Parameters.IntegralGain := LREAL#0.6666666666666667;
Parameters.ProportionalSetpointWeight := LREAL#1.0;
Parameters.Bias := LREAL#0.0;
Parameters.OutputMinimum := LREAL#-1.0e100;
Parameters.OutputMaximum := LREAL#1.0e100;
Parameters.RateMinimum := LREAL#-1.0e100;
Parameters.RateMaximum := LREAL#1.0e100;
Parameters.TrackingTime := LREAL#1.0;
State.Setpoint := LREAL#1.0;
State.ProcessValue := LREAL#1.0;
State.NominalOutput := LREAL#1.0;
State.SaturatedOutput := LREAL#1.0;
Controller.Configure(Parameters := Parameters);
Controller.Initialize(State := State);

Input.Setpoint := LREAL#3.0;
Input.ProcessValue := LREAL#1.0;
Input.CycleTime := LREAL#0.1;
Input.Mode := PIDMode#Auto;
Output := Controller.Update(Input := Input);
ASSERT_NEAR(EXPECTED := LREAL#2.4666666666666663, ACTUAL := Output, DELTA := LREAL#1.0e-12);

Parameters.IntegralGain := LREAL#0.0;
Parameters.Bias := LREAL#2.0;
Controller.Configure(Parameters := Parameters);
Input.ProcessValue := LREAL#2.9;
Output := Controller.Update(Input := Input);
ASSERT_NEAR(EXPECTED := LREAL#2.066666666666667, ACTUAL := Output, DELTA := LREAL#1.0e-12);

Parameters.IntegralGain := LREAL#0.6666666666666667;
Controller.Configure(Parameters := Parameters);
Input.Setpoint := LREAL#1.0;
Input.ProcessValue := LREAL#1.6;
Output := Controller.Update(Input := Input);
ASSERT_NEAR(EXPECTED := LREAL#1.56, ACTUAL := Output, DELTA := LREAL#1.0e-12);

Parameters.Bias := LREAL#0.0;
Parameters.RateMinimum := LREAL#-0.5;
Parameters.RateMaximum := LREAL#0.5;
LimitedController.Configure(Parameters := Parameters);
LimitedController.Initialize(State := State);
Input.Setpoint := LREAL#3.0;
Input.ProcessValue := LREAL#1.0;
Output := LimitedController.Update(Input := Input);
ASSERT_NEAR(EXPECTED := LREAL#1.05, ACTUAL := Output, DELTA := LREAL#1.0e-12);
END_TEST_PROGRAM

TEST_PROGRAM control_pid_replays_paper_example_3_setpoint_weighting
VAR
    FullWeight : PID;
    HalfWeight : PID;
    ZeroWeight : PID;
    Parameters : PIDParameters;
    State : PIDInitialState;
    Input : PIDInput;
    Output : LREAL;
END_VAR

Parameters.ProportionalGain := LREAL#0.6666666666666667;
Parameters.IntegralGain := LREAL#0.6666666666666667;
Parameters.ProportionalSetpointWeight := LREAL#1.0;
Parameters.OutputMinimum := LREAL#-1.0e100;
Parameters.OutputMaximum := LREAL#1.0e100;
Parameters.RateMinimum := LREAL#-1.0e100;
Parameters.RateMaximum := LREAL#1.0e100;
Parameters.TrackingTime := LREAL#1.0;
FullWeight.Configure(Parameters := Parameters);
FullWeight.Initialize(State := State);
Parameters.ProportionalSetpointWeight := LREAL#0.5;
HalfWeight.Configure(Parameters := Parameters);
HalfWeight.Initialize(State := State);
Parameters.ProportionalSetpointWeight := LREAL#0.0;
ZeroWeight.Configure(Parameters := Parameters);
ZeroWeight.Initialize(State := State);

Input.Setpoint := LREAL#3.0;
Input.CycleTime := LREAL#0.01;
Input.Mode := PIDMode#Auto;
Output := FullWeight.Update(Input := Input);
ASSERT_NEAR(EXPECTED := LREAL#2.02, ACTUAL := Output, DELTA := LREAL#1.0e-12);
Output := HalfWeight.Update(Input := Input);
ASSERT_NEAR(EXPECTED := LREAL#1.02, ACTUAL := Output, DELTA := LREAL#1.0e-12);
Output := ZeroWeight.Update(Input := Input);
ASSERT_NEAR(EXPECTED := LREAL#0.02, ACTUAL := Output, DELTA := LREAL#1.0e-12);

(* The same load disturbance changes the process-value term equally. *)
Input.ProcessValue := LREAL#1.0;
Output := FullWeight.Update(Input := Input);
ASSERT_NEAR(EXPECTED := LREAL#1.3666666666666667, ACTUAL := Output, DELTA := LREAL#1.0e-12);
Output := HalfWeight.Update(Input := Input);
ASSERT_NEAR(EXPECTED := LREAL#0.3666666666666667, ACTUAL := Output, DELTA := LREAL#1.0e-12);
Output := ZeroWeight.Update(Input := Input);
ASSERT_NEAR(EXPECTED := LREAL#-0.6333333333333333, ACTUAL := Output, DELTA := LREAL#1.0e-12);
END_TEST_PROGRAM

TEST_PROGRAM control_pid_replays_paper_example_4_feedforward_and_anti_windup
VAR
    Unconstrained : PID;
    Clamping : PID;
    BackCalculation : PID;
    Parameters : PIDParameters;
    State : PIDInitialState;
    Input : PIDInput;
    Output : LREAL;
END_VAR

Parameters.ProportionalGain := LREAL#2.727272727272727;
Parameters.IntegralGain := LREAL#0.9090909090909091;
Parameters.ProportionalSetpointWeight := LREAL#1.0;
Parameters.OutputMinimum := LREAL#-1.0e100;
Parameters.OutputMaximum := LREAL#1.0e100;
Parameters.RateMinimum := LREAL#-1.0e100;
Parameters.RateMaximum := LREAL#1.0e100;
Parameters.TrackingTime := LREAL#3.0;
Unconstrained.Configure(Parameters := Parameters);
Unconstrained.Initialize(State := State);
Parameters.OutputMinimum := LREAL#-3.5;
Parameters.OutputMaximum := LREAL#3.5;
Parameters.TrackingTime := LREAL#0.01;
Clamping.Configure(Parameters := Parameters);
Clamping.Initialize(State := State);
Parameters.TrackingTime := LREAL#3.0;
BackCalculation.Configure(Parameters := Parameters);
BackCalculation.Initialize(State := State);

Input.Setpoint := LREAL#4.5;
Input.CycleTime := LREAL#0.01;
Input.Mode := PIDMode#Auto;
Output := Unconstrained.Update(Input := Input);
ASSERT_NEAR(EXPECTED := LREAL#12.313636363636363, ACTUAL := Output, DELTA := LREAL#1.0e-11);
Output := Clamping.Update(Input := Input);
ASSERT_NEAR(EXPECTED := LREAL#3.5, ACTUAL := Output, DELTA := LREAL#1.0e-12);
Output := BackCalculation.Update(Input := Input);
ASSERT_NEAR(EXPECTED := LREAL#3.5, ACTUAL := Output, DELTA := LREAL#1.0e-12);

Input.Setpoint := LREAL#0.0;
Output := Clamping.Update(Input := Input);
ASSERT_NEAR(EXPECTED := LREAL#-3.5, ACTUAL := Output, DELTA := LREAL#1.0e-12);
Output := BackCalculation.Update(Input := Input);
ASSERT_NEAR(EXPECTED := LREAL#0.011530303030303557, ACTUAL := Output, DELTA := LREAL#1.0e-12);

Input.FeedForward := LREAL#-8.970083166928498;
Output := Unconstrained.Update(Input := Input);
ASSERT_NEAR(EXPECTED := LREAL#-8.929174076019407, ACTUAL := Output, DELTA := LREAL#1.0e-11);
Output := Clamping.Update(Input := Input);
ASSERT_NEAR(EXPECTED := LREAL#-3.5, ACTUAL := Output, DELTA := LREAL#1.0e-12);
Output := BackCalculation.Update(Input := Input);
ASSERT_NEAR(EXPECTED := LREAL#-3.5, ACTUAL := Output, DELTA := LREAL#1.0e-12);
END_TEST_PROGRAM

TEST_PROGRAM control_pid_replays_paper_example_5_measurement_filters
VAR
    SlowFirst : LowPass;
    SlowSecond : LowPass;
    FastFirst : LowPass;
    FastSecond : LowPass;
    Parameters : LowPassParameters;
    Output : LREAL;
END_VAR

Parameters.TimeConstant := LREAL#0.1;
Parameters.Order := FilterOrder#FirstOrder;
SlowFirst.Configure(Parameters := Parameters);
SlowFirst.Initialize(Input := LREAL#0.0);
Parameters.Order := FilterOrder#SecondOrder;
SlowSecond.Configure(Parameters := Parameters);
SlowSecond.Initialize(Input := LREAL#0.0);
Parameters.TimeConstant := LREAL#0.01;
Parameters.Order := FilterOrder#FirstOrder;
FastFirst.Configure(Parameters := Parameters);
FastFirst.Initialize(Input := LREAL#0.0);
Parameters.Order := FilterOrder#SecondOrder;
FastSecond.Configure(Parameters := Parameters);
FastSecond.Initialize(Input := LREAL#0.0);

(* These are selected released noisy measurements after the process delay. *)
Output := SlowFirst.Update(Input := LREAL#0.0775918043205658, CycleTime := LREAL#0.01);
Output := SlowFirst.Update(Input := LREAL#0.14700588752798377, CycleTime := LREAL#0.01);
Output := SlowFirst.Update(Input := LREAL#0.26877691165790607, CycleTime := LREAL#0.01);
ASSERT_NEAR(EXPECTED := LREAL#0.04431413638365756, ACTUAL := Output, DELTA := LREAL#1.0e-12);

Output := SlowSecond.Update(Input := LREAL#0.0775918043205658, CycleTime := LREAL#0.01);
Output := SlowSecond.Update(Input := LREAL#0.14700588752798377, CycleTime := LREAL#0.01);
Output := SlowSecond.Update(Input := LREAL#0.26877691165790607, CycleTime := LREAL#0.01);
ASSERT_NEAR(EXPECTED := LREAL#0.0065790126617539055, ACTUAL := Output, DELTA := LREAL#1.0e-12);

Output := FastFirst.Update(Input := LREAL#0.0775918043205658, CycleTime := LREAL#0.01);
Output := FastFirst.Update(Input := LREAL#0.14700588752798377, CycleTime := LREAL#0.01);
Output := FastFirst.Update(Input := LREAL#0.26877691165790607, CycleTime := LREAL#0.01);
ASSERT_NEAR(EXPECTED := LREAL#0.21760012383893867, ACTUAL := Output, DELTA := LREAL#1.0e-12);

Output := FastSecond.Update(Input := LREAL#0.0775918043205658, CycleTime := LREAL#0.01);
Output := FastSecond.Update(Input := LREAL#0.14700588752798377, CycleTime := LREAL#0.01);
Output := FastSecond.Update(Input := LREAL#0.26877691165790607, CycleTime := LREAL#0.01);
ASSERT_NEAR(EXPECTED := LREAL#0.17450878731114844, ACTUAL := Output, DELTA := LREAL#1.0e-12);
END_TEST_PROGRAM

TEST_PROGRAM control_pid_replays_paper_example_6_gain_scheduling_with_tracking
VAR
    LowController : PID;
    MiddleController : PID;
    HighController : PID;
    Parameters : PIDParameters;
    State : PIDInitialState;
    Input : PIDInput;
    TankArea : LREAL;
    OrificeArea : LREAL;
    Gravity : LREAL;
    Time1 : LREAL;
    Time2 : LREAL;
    Time3 : LREAL;
    Gain1 : LREAL;
    Gain2 : LREAL;
    Gain3 : LREAL;
    CommonTime : LREAL;
    InitialFlow : LREAL;
    LowOutput : LREAL;
    MiddleOutput : LREAL;
    HighOutput : LREAL;
    SelectedOutput : LREAL;
END_VAR

TankArea := LREAL#390.0;
OrificeArea := LREAL#2.15;
Gravity := LREAL#983.0;
Time1 := TankArea / OrificeArea * SQRT(LREAL#8.0 / Gravity);
Time2 := TankArea / OrificeArea * SQRT(LREAL#24.0 / Gravity);
Time3 := TankArea / OrificeArea * SQRT(LREAL#40.0 / Gravity);
Gain1 := Time1 / TankArea;
Gain2 := Time2 / TankArea;
Gain3 := Time3 / TankArea;
CommonTime := (Time1 + Time2 + Time3) / LREAL#3.0;
InitialFlow := OrificeArea * SQRT(LREAL#8.0 * Gravity);

Parameters.ProportionalGain := Time1 / (Gain1 * CommonTime);
Parameters.IntegralGain := Parameters.ProportionalGain / Time1;
Parameters.ProportionalSetpointWeight := LREAL#1.0;
Parameters.OutputMinimum := LREAL#-1.0e100;
Parameters.OutputMaximum := LREAL#1.0e100;
Parameters.RateMinimum := LREAL#-1.0e100;
Parameters.RateMaximum := LREAL#1.0e100;
Parameters.TrackingTime := Time1;
State.Setpoint := LREAL#4.0;
State.ProcessValue := LREAL#4.0;
State.NominalOutput := InitialFlow;
State.SaturatedOutput := InitialFlow;
LowController.Configure(Parameters := Parameters);
LowController.Initialize(State := State);
Parameters.ProportionalGain := Time2 / (Gain2 * CommonTime);
Parameters.IntegralGain := Parameters.ProportionalGain / Time2;
Parameters.TrackingTime := Time2;
MiddleController.Configure(Parameters := Parameters);
MiddleController.Initialize(State := State);
Parameters.ProportionalGain := Time3 / (Gain3 * CommonTime);
Parameters.IntegralGain := Parameters.ProportionalGain / Time3;
Parameters.TrackingTime := Time3;
HighController.Configure(Parameters := Parameters);
HighController.Initialize(State := State);

Input.Setpoint := LREAL#22.0;
Input.ProcessValue := LREAL#4.0;
Input.CycleTime := LREAL#0.01;
Input.Mode := PIDMode#Auto;
LowOutput := LowController.Update(Input := Input);
Input.Mode := PIDMode#Track;
Input.TrackingOutput := InitialFlow;
MiddleOutput := MiddleController.Update(Input := Input);
HighOutput := HighController.Update(Input := Input);
SelectedOutput := LowOutput;
ASSERT_NEAR(EXPECTED := LREAL#449.8616638937913, ACTUAL := SelectedOutput, DELTA := LREAL#1.0e-8);

Input.ProcessValue := LREAL#12.1;
Input.TrackingOutput := SelectedOutput;
Input.Mode := PIDMode#Track;
LowOutput := LowController.Update(Input := Input);
Input.Mode := PIDMode#Auto;
MiddleOutput := MiddleController.Update(Input := Input);
Input.Mode := PIDMode#Track;
HighOutput := HighController.Update(Input := Input);
SelectedOutput := MiddleOutput;
ASSERT_NEAR(EXPECTED := LREAL#333.2756344812609, ACTUAL := SelectedOutput, DELTA := LREAL#1.0e-8);

Input.ProcessValue := LREAL#20.1;
Input.TrackingOutput := SelectedOutput;
Input.Mode := PIDMode#Track;
LowOutput := LowController.Update(Input := Input);
MiddleOutput := MiddleController.Update(Input := Input);
Input.Mode := PIDMode#Auto;
HighOutput := HighController.Update(Input := Input);
SelectedOutput := HighOutput;
ASSERT_NEAR(EXPECTED := LREAL#218.20841899630443, ACTUAL := SelectedOutput, DELTA := LREAL#1.0e-8);
END_TEST_PROGRAM

TEST_PROGRAM control_pid_replays_paper_example_7_selector_with_tracking
VAR
    FirstController : PID;
    SecondController : PID;
    Parameters : PIDParameters;
    FirstState : PIDInitialState;
    SecondState : PIDInitialState;
    FirstInput : PIDInput;
    SecondInput : PIDInput;
    FirstOutput : LREAL;
    SecondOutput : LREAL;
    SelectedOutput : LREAL;
END_VAR

Parameters.ProportionalGain := LREAL#0.6666666666666667;
Parameters.IntegralGain := LREAL#0.6666666666666667;
Parameters.ProportionalSetpointWeight := LREAL#1.0;
Parameters.OutputMinimum := LREAL#-1.0e100;
Parameters.OutputMaximum := LREAL#1.0e100;
Parameters.RateMinimum := LREAL#-1.0e100;
Parameters.RateMaximum := LREAL#1.0e100;
Parameters.TrackingTime := LREAL#1.0;
FirstState.Setpoint := LREAL#0.3;
FirstState.ProcessValue := LREAL#0.3;
SecondState.Setpoint := LREAL#0.5;
SecondState.ProcessValue := LREAL#0.5;
FirstController.Configure(Parameters := Parameters);
FirstController.Initialize(State := FirstState);
SecondController.Configure(Parameters := Parameters);
SecondController.Initialize(State := SecondState);

FirstInput.Setpoint := LREAL#0.3;
FirstInput.ProcessValue := LREAL#0.2871535891077072;
FirstInput.CycleTime := LREAL#0.01;
FirstInput.Mode := PIDMode#Auto;
SecondInput.Setpoint := LREAL#0.5;
SecondInput.ProcessValue := LREAL#0.49502491687458405;
SecondInput.CycleTime := LREAL#0.01;
SecondInput.Mode := PIDMode#Track;
FirstOutput := FirstController.Update(Input := FirstInput);
SecondOutput := SecondController.Update(Input := SecondInput);
SelectedOutput := MIN(FirstOutput, SecondOutput);
ASSERT_NEAR(EXPECTED := LREAL#0.003349889304446737, ACTUAL := SelectedOutput, DELTA := LREAL#1.0e-12);

FirstInput.ProcessValue := LREAL#0.2785272123191362;
FirstInput.TrackingOutput := SelectedOutput;
FirstInput.Mode := PIDMode#Track;
SecondInput.ProcessValue := LREAL#0.5;
SecondInput.TrackingOutput := SelectedOutput;
SecondInput.Mode := PIDMode#Auto;
FirstOutput := FirstController.Update(Input := FirstInput);
SecondOutput := SecondController.Update(Input := SecondInput);
SelectedOutput := MIN(FirstOutput, SecondOutput);
ASSERT_NEAR(EXPECTED := LREAL#0.00003316722083610609, ACTUAL := SelectedOutput, DELTA := LREAL#1.0e-12);

FirstInput.ProcessValue := LREAL#0.2682;
FirstInput.TrackingOutput := SelectedOutput;
SecondInput.ProcessValue := LREAL#0.447019;
SecondInput.TrackingOutput := SelectedOutput;
FirstOutput := FirstController.Update(Input := FirstInput);
SecondOutput := SecondController.Update(Input := SecondInput);
SelectedOutput := MIN(FirstOutput, SecondOutput);
ASSERT_NEAR(EXPECTED := LREAL#0.0071299754335935675, ACTUAL := SelectedOutput, DELTA := LREAL#1.0e-12);
END_TEST_PROGRAM

(* ---- term_tests.st ---- *)
USING Control;

TEST_PROGRAM control_pid_feedforward_is_positional_incremental_and_manual_history_aware
VAR
    PositionalController : PID;
    IncrementalController : PID;
    ManualController : PID;
    Parameters : PIDParameters;
    InitialState : PIDInitialState;
    Input : PIDInput;
    Output : LREAL;
END_VAR

Parameters.OutputMinimum := LREAL#-100.0;
Parameters.OutputMaximum := LREAL#100.0;
Parameters.RateMinimum := LREAL#-1000.0;
Parameters.RateMaximum := LREAL#1000.0;
Parameters.TrackingTime := LREAL#1.0;

PositionalController.Configure(Parameters := Parameters);
PositionalController.Initialize(State := InitialState);
Input.FeedForward := LREAL#2.0;
Input.CycleTime := LREAL#0.1;
Output := PositionalController.Update(Input := Input);
ASSERT_NEAR(EXPECTED := LREAL#2.0, ACTUAL := Output, DELTA := LREAL#2.0e-12);

Parameters.IntegralGain := LREAL#1.0;
InitialState.FeedForward := LREAL#1.0;
InitialState.NominalOutput := LREAL#10.0;
InitialState.SaturatedOutput := LREAL#10.0;
IncrementalController.Configure(Parameters := Parameters);
IncrementalController.Initialize(State := InitialState);
Input.FeedForward := LREAL#3.0;
Output := IncrementalController.Update(Input := Input);
ASSERT_NEAR(EXPECTED := LREAL#12.0, ACTUAL := Output, DELTA := LREAL#12.0e-12);

InitialState.FeedForward := LREAL#1.0;
InitialState.NominalOutput := LREAL#0.0;
InitialState.SaturatedOutput := LREAL#0.0;
ManualController.Configure(Parameters := Parameters);
ManualController.Initialize(State := InitialState);
Input.FeedForward := LREAL#5.0;
Input.ManualOutput := LREAL#7.0;
Input.Mode := PIDMode#Manual;
Output := ManualController.Update(Input := Input);
ASSERT_NEAR(EXPECTED := LREAL#7.0, ACTUAL := Output, DELTA := LREAL#7.0e-12);
Input.Mode := PIDMode#Auto;
Output := ManualController.Update(Input := Input);
ASSERT_NEAR(EXPECTED := LREAL#7.0, ACTUAL := Output, DELTA := LREAL#7.0e-12);
END_TEST_PROGRAM

TEST_PROGRAM control_pid_setpoint_weights_affect_only_their_paper_terms
VAR
    ControllerA : PID;
    ControllerB : PID;
    Parameters : PIDParameters;
    InitialState : PIDInitialState;
    Input : PIDInput;
    Output : LREAL;
END_VAR

Parameters.ProportionalGain := LREAL#2.0;
Parameters.IntegralGain := LREAL#1.0;
Parameters.ProportionalSetpointWeight := LREAL#0.25;
Parameters.OutputMinimum := LREAL#-100.0;
Parameters.OutputMaximum := LREAL#100.0;
Parameters.RateMinimum := LREAL#-1000.0;
Parameters.RateMaximum := LREAL#1000.0;
Parameters.TrackingTime := LREAL#1.0;
ControllerA.Configure(Parameters := Parameters);
ControllerA.Initialize(State := InitialState);
Input.Setpoint := LREAL#2.0;
Input.ProcessValue := LREAL#0.5;
Input.CycleTime := LREAL#0.1;
Output := ControllerA.Update(Input := Input);
ASSERT_NEAR(EXPECTED := LREAL#0.15, ACTUAL := Output, DELTA := LREAL#1.0e-12);

Parameters.ProportionalSetpointWeight := LREAL#0.75;
ControllerB.Configure(Parameters := Parameters);
ControllerB.Initialize(State := InitialState);
Output := ControllerB.Update(Input := Input);
ASSERT_NEAR(EXPECTED := LREAL#2.15, ACTUAL := Output, DELTA := LREAL#2.15e-12);

Parameters.IntegralGain := LREAL#0.0;
Parameters.ProportionalSetpointWeight := LREAL#0.0;
ControllerA.Configure(Parameters := Parameters);
ControllerA.Initialize(State := InitialState);
Output := ControllerA.Update(Input := Input);
ASSERT_NEAR(EXPECTED := LREAL#3.0, ACTUAL := Output, DELTA := LREAL#3.0e-12);

Parameters.ProportionalGain := LREAL#0.0;
Parameters.DerivativeGain := LREAL#0.5;
Parameters.DerivativeSetpointWeight := LREAL#0.25;
ControllerA.Configure(Parameters := Parameters);
ControllerA.Initialize(State := InitialState);
Output := ControllerA.Update(Input := Input);
ASSERT_NEAR(EXPECTED := LREAL#0.0, ACTUAL := Output, DELTA := LREAL#1.0e-12);

Parameters.DerivativeSetpointWeight := LREAL#0.0;
ControllerB.Configure(Parameters := Parameters);
ControllerB.Initialize(State := InitialState);
Output := ControllerB.Update(Input := Input);
ASSERT_NEAR(EXPECTED := LREAL#-2.5, ACTUAL := Output, DELTA := LREAL#2.5e-12);

Parameters.IntegralGain := LREAL#1.0;
Parameters.DerivativeSetpointWeight := LREAL#0.25;
ControllerA.Configure(Parameters := Parameters);
ControllerA.Initialize(State := InitialState);
Output := ControllerA.Update(Input := Input);
ASSERT_NEAR(EXPECTED := LREAL#0.15, ACTUAL := Output, DELTA := LREAL#1.0e-12);

Parameters.DerivativeSetpointWeight := LREAL#0.0;
ControllerB.Configure(Parameters := Parameters);
ControllerB.Initialize(State := InitialState);
Output := ControllerB.Update(Input := Input);
ASSERT_NEAR(EXPECTED := LREAL#-2.35, ACTUAL := Output, DELTA := LREAL#2.35e-12);
END_TEST_PROGRAM

(* ---- tests.st ---- *)
TEST_PROGRAM control_pid_positional_pd_uses_actual_cycle_time
VAR
    Controller : Control.PID;
    Parameters : Control.PIDParameters;
    InitialState : Control.PIDInitialState;
    Input : Control.PIDInput;
    Output : LREAL;
END_VAR

Parameters.ProportionalGain := LREAL#2.0;
Parameters.IntegralGain := LREAL#0.0;
Parameters.DerivativeGain := LREAL#0.5;
Parameters.ProportionalSetpointWeight := LREAL#0.0;
Parameters.DerivativeSetpointWeight := LREAL#0.25;
Parameters.Bias := LREAL#1.0;
Parameters.OutputMinimum := LREAL#-100.0;
Parameters.OutputMaximum := LREAL#100.0;
Parameters.RateMinimum := LREAL#-1000.0;
Parameters.RateMaximum := LREAL#1000.0;
Parameters.TrackingTime := LREAL#1.0;

Controller.Configure(Parameters := Parameters);
Controller.Initialize(State := InitialState);

Input.Setpoint := LREAL#1.0;
Input.ProcessValue := LREAL#0.2;
Input.FeedForward := LREAL#0.3;
Input.CycleTime := LREAL#0.1;
Output := Controller.Update(Input := Input);
ASSERT_NEAR(EXPECTED := LREAL#3.15, ACTUAL := Output, DELTA := LREAL#3.15e-12);

Input.ProcessValue := LREAL#0.4;
Input.CycleTime := LREAL#0.2;
Output := Controller.Update(Input := Input);
ASSERT_NEAR(EXPECTED := LREAL#2.0, ACTUAL := Output, DELTA := LREAL#2.0e-12);
END_TEST_PROGRAM

TEST_PROGRAM control_pid_switches_forms_without_resetting_nominal_history
VAR
    Controller : Control.PID;
    Parameters : Control.PIDParameters;
    InitialState : Control.PIDInitialState;
    Input : Control.PIDInput;
    Output : LREAL;
END_VAR

Parameters.ProportionalGain := LREAL#2.0;
Parameters.IntegralGain := LREAL#0.5;
Parameters.ProportionalSetpointWeight := LREAL#0.5;
Parameters.Bias := LREAL#1.0;
Parameters.OutputMinimum := LREAL#-100.0;
Parameters.OutputMaximum := LREAL#100.0;
Parameters.RateMinimum := LREAL#-1000.0;
Parameters.RateMaximum := LREAL#1000.0;
Parameters.TrackingTime := LREAL#1.0;
Controller.Configure(Parameters := Parameters);
Controller.Initialize(State := InitialState);

Input.Setpoint := LREAL#1.0;
Input.CycleTime := LREAL#0.1;
Output := Controller.Update(Input := Input);
ASSERT_NEAR(EXPECTED := LREAL#1.05, ACTUAL := Output, DELTA := LREAL#1.05e-12);

Parameters.IntegralGain := LREAL#0.0;
Controller.Configure(Parameters := Parameters);
Output := Controller.Update(Input := Input);
ASSERT_NEAR(EXPECTED := LREAL#3.0, ACTUAL := Output, DELTA := LREAL#3.0e-12);

Parameters.IntegralGain := LREAL#0.5;
Controller.Configure(Parameters := Parameters);
Output := Controller.Update(Input := Input);
ASSERT_NEAR(EXPECTED := LREAL#3.05, ACTUAL := Output, DELTA := LREAL#3.05e-12);

Parameters.ProportionalGain := LREAL#4.0;
Controller.Configure(Parameters := Parameters);
Output := Controller.Update(Input := Input);
ASSERT_NEAR(EXPECTED := LREAL#3.10, ACTUAL := Output, DELTA := LREAL#3.10e-12);
END_TEST_PROGRAM

TEST_PROGRAM control_pid_incremental_pi_and_pid_use_signal_differences
VAR
    PidController : Control.PID;
    PiController : Control.PID;
    Parameters : Control.PIDParameters;
    InitialState : Control.PIDInitialState;
    Input : Control.PIDInput;
    Output : LREAL;
END_VAR

Parameters.ProportionalGain := LREAL#2.0;
Parameters.IntegralGain := LREAL#0.5;
Parameters.DerivativeGain := LREAL#0.1;
Parameters.ProportionalSetpointWeight := LREAL#0.5;
Parameters.DerivativeSetpointWeight := LREAL#0.0;
Parameters.OutputMinimum := LREAL#-100.0;
Parameters.OutputMaximum := LREAL#100.0;
Parameters.RateMinimum := LREAL#-1000.0;
Parameters.RateMaximum := LREAL#1000.0;
Parameters.TrackingTime := LREAL#1.0;

PidController.Configure(Parameters := Parameters);
PidController.Initialize(State := InitialState);

Input.Setpoint := LREAL#1.0;
Input.ProcessValue := LREAL#0.0;
Input.FeedForward := LREAL#0.2;
Input.CycleTime := LREAL#0.1;
Output := PidController.Update(Input := Input);
ASSERT_NEAR(EXPECTED := LREAL#1.25, ACTUAL := Output, DELTA := LREAL#1.25e-12);

Input.ProcessValue := LREAL#0.2;
Input.FeedForward := LREAL#0.3;
Output := PidController.Update(Input := Input);
ASSERT_NEAR(EXPECTED := LREAL#0.79, ACTUAL := Output, DELTA := LREAL#1.0e-12);

Parameters.DerivativeGain := LREAL#0.0;
PiController.Configure(Parameters := Parameters);
PiController.Initialize(State := InitialState);

Input.ProcessValue := LREAL#0.0;
Input.FeedForward := LREAL#0.2;
Output := PiController.Update(Input := Input);
ASSERT_NEAR(EXPECTED := LREAL#1.25, ACTUAL := Output, DELTA := LREAL#1.25e-12);

Input.ProcessValue := LREAL#0.2;
Input.FeedForward := LREAL#0.3;
Output := PiController.Update(Input := Input);
ASSERT_NEAR(EXPECTED := LREAL#0.99, ACTUAL := Output, DELTA := LREAL#1.0e-12);
END_TEST_PROGRAM
